{attribute 'Tc2GvlVarNames'}
VAR_GLOBAL
(* Inputs / Eingänge *)
	binGr02LightCurtainOK					AT %I*:BOOL;													(*) 	Light curtain ok / Freigabe Lichtschranke i.o *)

	binGr02PushBtnStart						AT %I*:BOOL;													(*) 	Push button "Start" / Taste "Start" *)
	binGr02PushBtnStop						AT %I*:BOOL;													(*) 	Push button "Stop" / Taste "Stop" *)

	(* Outputs / Ausgänge *)
	boutGr02ConfLightCurtain				AT %Q*:BOOL;													(*) 	Confirm light Curtain / Quitt Lichtschrank *)

	boutGr02BulbBtnStart					AT %Q*:BOOL;													(*) 	Signal button bulb "start" / Signallampe "Start" *)
	boutGr02BulbBtnStop						AT %Q*:BOOL;													(*) 	Signal button bulb "stop" / Signallampe "Stop" *)

END_VAR

(* stored: Version 1.1.0.1, ProductVersion 3.1.4024.15
   GVL GVL_Gr02IO: Id {f045defe-70af-469a-a92d-ee44c7ef8f87} *)
